(* IEC 61131-3 sources: iFA_git_test/GIT test/PLC_1/Programs, 4 files *)

(* ---- DefaultVariableTable.st ---- *)
(*NodeCRC64:15794442468608431415, FileCRC64:15794442468608431415*)
VAR_GLOBAL
END_VAR
(*{"Version":"1.0.0.0","Path":"Default_variable_table","ObjectType":"Global"}*)
END_VAR_GLOBAL

(* ---- FB_Example.st ---- *)
(*NodeCRC64:9907401017642776752, FileCRC64:9907401017642776752*)
FUNCTION_BLOCK FB_Example
VAR_INPUT
END_VAR
VAR_OUTPUT
END_VAR
VAR
END_VAR
Body

EndBody
(*{"Version":"1.0.0.0","Path":"FB_Example","ObjectType":"FunctionBlock"}*)
END_FUNCTION_BLOCK

(* ---- Main.st ---- *)
(*NodeCRC64:8187142076338617645, FileCRC64:8187142076338617645*)
PROGRAM Main
VAR
    liCounter : LINT;
    liCounter2 : LINT;
END_VAR
Body
liCounter := liCounter + 1;
EndBody
(*{"Version":"1.0.0.0","Path":"Main","ObjectType":"Program"}*)
END_PROGRAM

(* ---- TestFBFromGIT.st ---- *)
PROGRAM TestFBFromGIT
VAR
    liCounter : LINT;
    liCounter2 : LINT;
END_VAR
Body
liCounter := liCounter + 1;
EndBody
(*{"Version":"1.0.0.0","Path":"TestFBFromGIT","ObjectType":"Program"}*)
END_PROGRAM
